(* IEC 61131-3 sources: sis-interlock-demo/pytests/golden/mini/src/POUs/Generated/FB_SisApp, 1 file *)

(* ---- FB_SisApp.decl.st ---- *)
// AUTO-GENERATED by cemgen 1.0.0 — не редактировать: правьте матрицу и запустите
//   python -m cemgen generate <файл матрицы .csv или .xlsx>
// Матрица: TEST-U301-CEM, объект U-301, ревизия 1 от 2026-10-16, SHA-256 сетки 9067fda96ae55e67
// Назначение: привязка ПАЗ объекта U-301 к образу ввода-вывода: токи 4–20 мА → инж. ед. и
//             достоверность по NE 43, дискретные входы и контроль линии → группы голосования по
//             причинам; вызов FB_SisUnit с конфигурацией GVL_SisCfg; разрешения следствий → выходы
//             xQ*.
// Автор:      pytest; код — генератор cemgen
// Версия:     1.0.0
// Документ:   docs/DESIGN.md, раздел «10. Генератор cemgen»; docs/cause_effect_matrix.md
// ВНИМАНИЕ:   код демонстрационный и не предназначен для систем безопасности. Реальная ПАЗ требует
//             определения SIL, сертифицированных аппаратных и программных средств и валидации по
//             ГОСТ Р МЭК 61511.
FUNCTION_BLOCK FB_SisApp
VAR_INPUT
    itfTime : PL.I_TimeSource;      // 0 — системное время
    itfLog  : I_SisEventSink;       // 0 — без журнала
END_VAR
VAR_IN_OUT
    stIo  : ST_SisIo;               // входы читает, выходы xQ* пишет
    stCmd : ST_SisCmd;              // команды HMI
END_VAR
VAR_OUTPUT
    xTripped   : BOOL := TRUE;                                          // сработало хотя бы одно следствие
    stCemSts   : ST_CauseEffectSts;                                     // состояние матрицы
    astVoteSts : ARRAY[1..GVL_Const.SIS_CAUSES_MAX] OF ST_VotingSts;   // состояние групп голосования
END_VAR
VAR
    fbUnit : FB_SisUnit;                                                // общий узел ПАЗ
    astIn  : ARRAY[1..GVL_Const.SIS_CAUSES_MAX] OF ST_VoteIn;       // входы групп по причинам
END_VAR
